// TIA Portal V21 export
DATA_BLOCK "Issue221_unit_plain"   // DB
{ S7_Optimized_Access := 'TRUE' }
// stored: AutoNumber true
BEGIN
END_DATA_BLOCK
